// Mitsubishi GX Works2 project: Task_4_Ex   PLC: FX3G

PROGRAM MAIN
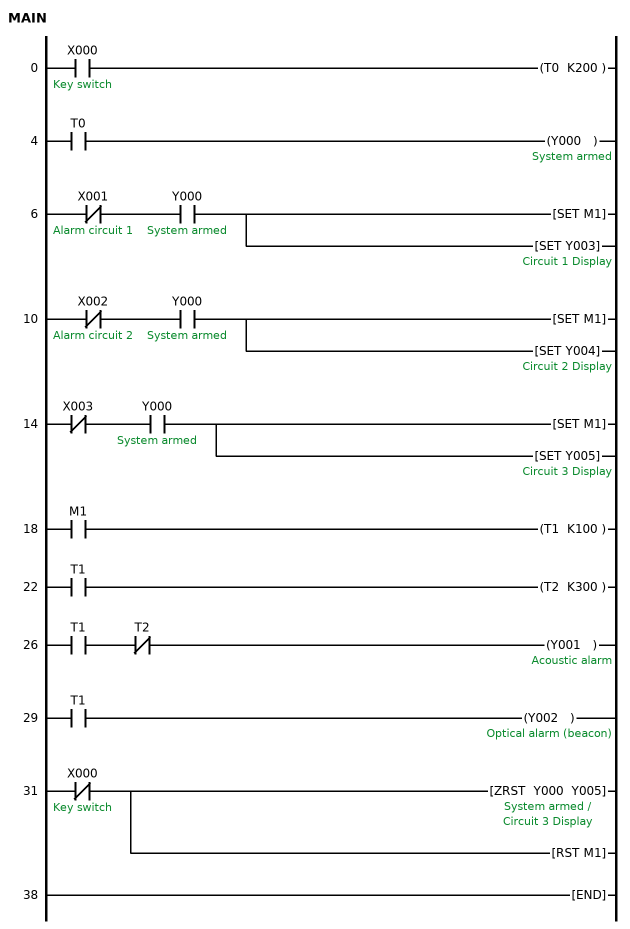
0     LD      X000  ; Key switch
      OUT     T0 K200
4     LD      T0
      OUT     Y000  ; System armed
6     LDI     X001  ; Alarm circuit 1
      AND     Y000  ; System armed
      SET     M1
      SET     Y003  ; Circuit 1 Display
10    LDI     X002  ; Alarm circuit 2
      AND     Y000  ; System armed
      SET     M1
      SET     Y004  ; Circuit 2 Display
14    LDI     X003
      AND     Y000  ; System armed
      SET     M1
      SET     Y005  ; Circuit 3 Display
18    LD      M1
      OUT     T1 K100
22    LD      T1
      OUT     T2 K300
26    LD      T1
      ANI     T2
      OUT     Y001  ; Acoustic alarm
29    LD      T1
      OUT     Y002  ; Optical alarm (beacon)
31    LDI     X000  ; Key switch
      ZRST    Y000 Y005
      RST     M1
38    END
END_PROGRAM
